DATA_BLOCK "GDB_GRAPH_PressDemoAuto"
{ S7_Optimized_Access := 'TRUE' }
VERSION : 0.1
NON_RETAIN
"FB_GRAPH_PressDemoAuto"
BEGIN
END_DATA_BLOCK
